Fanuc KAREL source: KT00580.KL

PROGRAM KT00580
%NOLOCKGROUP
VAR
  V1: VECTOR
  I2: INTEGER
  OUT: VECTOR
BEGIN
  V1.X = 1.0
    I2 = 3
  OUT = V1 / I2
END KT00580
